(* IEC 61131-3 sources: STAR-PLC-Agent/results/raw/four_group_20261114/star_deepseek_v4/PUB019/generation/sim_00, 1 file *)

(* ---- test_program.st ---- *)
PROGRAM PLC_PRG
VAR
 BenchStep : UDINT := 0;
 BenchCalls : UDINT := 0;
 BenchDone : BOOL := FALSE;
 BenchUut0 : FB_Task;
 BenchUut1 : FB_Task;
 TraceIn_ManualMode : ARRAY[0..12] OF BOOL;
 TraceIn_SingleStepMode : ARRAY[0..12] OF BOOL;
 TraceIn_SingleCycleMode : ARRAY[0..12] OF BOOL;
 TraceIn_ContinuousMode : ARRAY[0..12] OF BOOL;
 TraceIn_EmergencyStop : ARRAY[0..12] OF BOOL;
 TraceIn_Start : ARRAY[0..12] OF BOOL;
 TraceIn_DownButton : ARRAY[0..12] OF BOOL;
 TraceIn_UpButton : ARRAY[0..12] OF BOOL;
 TraceIn_LeftButton : ARRAY[0..12] OF BOOL;
 TraceIn_RightButton : ARRAY[0..12] OF BOOL;
 TraceIn_GripButton : ARRAY[0..12] OF BOOL;
 TraceIn_ReleaseButton : ARRAY[0..12] OF BOOL;
 TraceIn_DownLimitSwitch : ARRAY[0..12] OF BOOL;
 TraceIn_UpLimitSwitch : ARRAY[0..12] OF BOOL;
 TraceIn_LeftLimitSwitch : ARRAY[0..12] OF BOOL;
 TraceIn_RightLimitSwitch : ARRAY[0..12] OF BOOL;
 TraceIn_GripLimitSwitch : ARRAY[0..12] OF BOOL;
 TraceIn_ReleaseLimitSwitch : ARRAY[0..12] OF BOOL;
 TraceOut_MoveDown : ARRAY[0..12] OF BOOL;
 TraceOut_MoveUp : ARRAY[0..12] OF BOOL;
 TraceOut_MoveLeft : ARRAY[0..12] OF BOOL;
 TraceOut_MoveRight : ARRAY[0..12] OF BOOL;
 TraceOut_ActivateGrip : ARRAY[0..12] OF BOOL;
 TraceOut_ActivateRelease : ARRAY[0..12] OF BOOL;
END_VAR

IF NOT BenchDone THEN
 CASE BenchStep OF
 0:
   BenchUut0.ManualMode := TRUE;
   BenchUut0.SingleStepMode := FALSE;
   BenchUut0.SingleCycleMode := FALSE;
   BenchUut0.ContinuousMode := FALSE;
   BenchUut0.EmergencyStop := TRUE;
   BenchUut0.Start := FALSE;
   BenchUut0.DownButton := TRUE;
   BenchUut0.UpButton := FALSE;
   BenchUut0.LeftButton := FALSE;
   BenchUut0.RightButton := FALSE;
   BenchUut0.GripButton := FALSE;
   BenchUut0.ReleaseButton := FALSE;
   BenchUut0.DownLimitSwitch := FALSE;
   BenchUut0.UpLimitSwitch := TRUE;
   BenchUut0.LeftLimitSwitch := TRUE;
   BenchUut0.RightLimitSwitch := FALSE;
   BenchUut0.GripLimitSwitch := FALSE;
   BenchUut0.ReleaseLimitSwitch := FALSE;
   TraceIn_ManualMode[0] := BenchUut0.ManualMode;
   TraceIn_SingleStepMode[0] := BenchUut0.SingleStepMode;
   TraceIn_SingleCycleMode[0] := BenchUut0.SingleCycleMode;
   TraceIn_ContinuousMode[0] := BenchUut0.ContinuousMode;
   TraceIn_EmergencyStop[0] := BenchUut0.EmergencyStop;
   TraceIn_Start[0] := BenchUut0.Start;
   TraceIn_DownButton[0] := BenchUut0.DownButton;
   TraceIn_UpButton[0] := BenchUut0.UpButton;
   TraceIn_LeftButton[0] := BenchUut0.LeftButton;
   TraceIn_RightButton[0] := BenchUut0.RightButton;
   TraceIn_GripButton[0] := BenchUut0.GripButton;
   TraceIn_ReleaseButton[0] := BenchUut0.ReleaseButton;
   TraceIn_DownLimitSwitch[0] := BenchUut0.DownLimitSwitch;
   TraceIn_UpLimitSwitch[0] := BenchUut0.UpLimitSwitch;
   TraceIn_LeftLimitSwitch[0] := BenchUut0.LeftLimitSwitch;
   TraceIn_RightLimitSwitch[0] := BenchUut0.RightLimitSwitch;
   TraceIn_GripLimitSwitch[0] := BenchUut0.GripLimitSwitch;
   TraceIn_ReleaseLimitSwitch[0] := BenchUut0.ReleaseLimitSwitch;
   BenchUut0();
   TraceOut_MoveDown[0] := BenchUut0.MoveDown;
   TraceOut_MoveUp[0] := BenchUut0.MoveUp;
   TraceOut_MoveLeft[0] := BenchUut0.MoveLeft;
   TraceOut_MoveRight[0] := BenchUut0.MoveRight;
   TraceOut_ActivateGrip[0] := BenchUut0.ActivateGrip;
   TraceOut_ActivateRelease[0] := BenchUut0.ActivateRelease;
   BenchCalls := BenchCalls + 1;
 1:
   BenchUut0.ManualMode := TRUE;
   BenchUut0.SingleStepMode := FALSE;
   BenchUut0.SingleCycleMode := FALSE;
   BenchUut0.ContinuousMode := FALSE;
   BenchUut0.EmergencyStop := TRUE;
   BenchUut0.Start := FALSE;
   BenchUut0.DownButton := TRUE;
   BenchUut0.UpButton := FALSE;
   BenchUut0.LeftButton := FALSE;
   BenchUut0.RightButton := FALSE;
   BenchUut0.GripButton := FALSE;
   BenchUut0.ReleaseButton := FALSE;
   BenchUut0.DownLimitSwitch := TRUE;
   BenchUut0.UpLimitSwitch := FALSE;
   BenchUut0.LeftLimitSwitch := TRUE;
   BenchUut0.RightLimitSwitch := FALSE;
   BenchUut0.GripLimitSwitch := FALSE;
   BenchUut0.ReleaseLimitSwitch := FALSE;
   TraceIn_ManualMode[1] := BenchUut0.ManualMode;
   TraceIn_SingleStepMode[1] := BenchUut0.SingleStepMode;
   TraceIn_SingleCycleMode[1] := BenchUut0.SingleCycleMode;
   TraceIn_ContinuousMode[1] := BenchUut0.ContinuousMode;
   TraceIn_EmergencyStop[1] := BenchUut0.EmergencyStop;
   TraceIn_Start[1] := BenchUut0.Start;
   TraceIn_DownButton[1] := BenchUut0.DownButton;
   TraceIn_UpButton[1] := BenchUut0.UpButton;
   TraceIn_LeftButton[1] := BenchUut0.LeftButton;
   TraceIn_RightButton[1] := BenchUut0.RightButton;
   TraceIn_GripButton[1] := BenchUut0.GripButton;
   TraceIn_ReleaseButton[1] := BenchUut0.ReleaseButton;
   TraceIn_DownLimitSwitch[1] := BenchUut0.DownLimitSwitch;
   TraceIn_UpLimitSwitch[1] := BenchUut0.UpLimitSwitch;
   TraceIn_LeftLimitSwitch[1] := BenchUut0.LeftLimitSwitch;
   TraceIn_RightLimitSwitch[1] := BenchUut0.RightLimitSwitch;
   TraceIn_GripLimitSwitch[1] := BenchUut0.GripLimitSwitch;
   TraceIn_ReleaseLimitSwitch[1] := BenchUut0.ReleaseLimitSwitch;
   BenchUut0();
   TraceOut_MoveDown[1] := BenchUut0.MoveDown;
   TraceOut_MoveUp[1] := BenchUut0.MoveUp;
   TraceOut_MoveLeft[1] := BenchUut0.MoveLeft;
   TraceOut_MoveRight[1] := BenchUut0.MoveRight;
   TraceOut_ActivateGrip[1] := BenchUut0.ActivateGrip;
   TraceOut_ActivateRelease[1] := BenchUut0.ActivateRelease;
   BenchCalls := BenchCalls + 1;
 2:
   BenchUut0.ManualMode := TRUE;
   BenchUut0.SingleStepMode := FALSE;
   BenchUut0.SingleCycleMode := FALSE;
   BenchUut0.ContinuousMode := FALSE;
   BenchUut0.EmergencyStop := FALSE;
   BenchUut0.Start := FALSE;
   BenchUut0.DownButton := TRUE;
   BenchUut0.UpButton := FALSE;
   BenchUut0.LeftButton := FALSE;
   BenchUut0.RightButton := FALSE;
   BenchUut0.GripButton := FALSE;
   BenchUut0.ReleaseButton := FALSE;
   BenchUut0.DownLimitSwitch := FALSE;
   BenchUut0.UpLimitSwitch := TRUE;
   BenchUut0.LeftLimitSwitch := TRUE;
   BenchUut0.RightLimitSwitch := FALSE;
   BenchUut0.GripLimitSwitch := FALSE;
   BenchUut0.ReleaseLimitSwitch := FALSE;
   TraceIn_ManualMode[2] := BenchUut0.ManualMode;
   TraceIn_SingleStepMode[2] := BenchUut0.SingleStepMode;
   TraceIn_SingleCycleMode[2] := BenchUut0.SingleCycleMode;
   TraceIn_ContinuousMode[2] := BenchUut0.ContinuousMode;
   TraceIn_EmergencyStop[2] := BenchUut0.EmergencyStop;
   TraceIn_Start[2] := BenchUut0.Start;
   TraceIn_DownButton[2] := BenchUut0.DownButton;
   TraceIn_UpButton[2] := BenchUut0.UpButton;
   TraceIn_LeftButton[2] := BenchUut0.LeftButton;
   TraceIn_RightButton[2] := BenchUut0.RightButton;
   TraceIn_GripButton[2] := BenchUut0.GripButton;
   TraceIn_ReleaseButton[2] := BenchUut0.ReleaseButton;
   TraceIn_DownLimitSwitch[2] := BenchUut0.DownLimitSwitch;
   TraceIn_UpLimitSwitch[2] := BenchUut0.UpLimitSwitch;
   TraceIn_LeftLimitSwitch[2] := BenchUut0.LeftLimitSwitch;
   TraceIn_RightLimitSwitch[2] := BenchUut0.RightLimitSwitch;
   TraceIn_GripLimitSwitch[2] := BenchUut0.GripLimitSwitch;
   TraceIn_ReleaseLimitSwitch[2] := BenchUut0.ReleaseLimitSwitch;
   BenchUut0();
   TraceOut_MoveDown[2] := BenchUut0.MoveDown;
   TraceOut_MoveUp[2] := BenchUut0.MoveUp;
   TraceOut_MoveLeft[2] := BenchUut0.MoveLeft;
   TraceOut_MoveRight[2] := BenchUut0.MoveRight;
   TraceOut_ActivateGrip[2] := BenchUut0.ActivateGrip;
   TraceOut_ActivateRelease[2] := BenchUut0.ActivateRelease;
   BenchCalls := BenchCalls + 1;
 3:
   BenchUut0.ManualMode := TRUE;
   BenchUut0.SingleStepMode := FALSE;
   BenchUut0.SingleCycleMode := FALSE;
   BenchUut0.ContinuousMode := FALSE;
   BenchUut0.EmergencyStop := TRUE;
   BenchUut0.Start := FALSE;
   BenchUut0.DownButton := TRUE;
   BenchUut0.UpButton := FALSE;
   BenchUut0.LeftButton := FALSE;
   BenchUut0.RightButton := FALSE;
   BenchUut0.GripButton := FALSE;
   BenchUut0.ReleaseButton := FALSE;
   BenchUut0.DownLimitSwitch := FALSE;
   BenchUut0.UpLimitSwitch := TRUE;
   BenchUut0.LeftLimitSwitch := TRUE;
   BenchUut0.RightLimitSwitch := FALSE;
   BenchUut0.GripLimitSwitch := FALSE;
   BenchUut0.ReleaseLimitSwitch := FALSE;
   TraceIn_ManualMode[3] := BenchUut0.ManualMode;
   TraceIn_SingleStepMode[3] := BenchUut0.SingleStepMode;
   TraceIn_SingleCycleMode[3] := BenchUut0.SingleCycleMode;
   TraceIn_ContinuousMode[3] := BenchUut0.ContinuousMode;
   TraceIn_EmergencyStop[3] := BenchUut0.EmergencyStop;
   TraceIn_Start[3] := BenchUut0.Start;
   TraceIn_DownButton[3] := BenchUut0.DownButton;
   TraceIn_UpButton[3] := BenchUut0.UpButton;
   TraceIn_LeftButton[3] := BenchUut0.LeftButton;
   TraceIn_RightButton[3] := BenchUut0.RightButton;
   TraceIn_GripButton[3] := BenchUut0.GripButton;
   TraceIn_ReleaseButton[3] := BenchUut0.ReleaseButton;
   TraceIn_DownLimitSwitch[3] := BenchUut0.DownLimitSwitch;
   TraceIn_UpLimitSwitch[3] := BenchUut0.UpLimitSwitch;
   TraceIn_LeftLimitSwitch[3] := BenchUut0.LeftLimitSwitch;
   TraceIn_RightLimitSwitch[3] := BenchUut0.RightLimitSwitch;
   TraceIn_GripLimitSwitch[3] := BenchUut0.GripLimitSwitch;
   TraceIn_ReleaseLimitSwitch[3] := BenchUut0.ReleaseLimitSwitch;
   BenchUut0();
   TraceOut_MoveDown[3] := BenchUut0.MoveDown;
   TraceOut_MoveUp[3] := BenchUut0.MoveUp;
   TraceOut_MoveLeft[3] := BenchUut0.MoveLeft;
   TraceOut_MoveRight[3] := BenchUut0.MoveRight;
   TraceOut_ActivateGrip[3] := BenchUut0.ActivateGrip;
   TraceOut_ActivateRelease[3] := BenchUut0.ActivateRelease;
   BenchCalls := BenchCalls + 1;
 4:
   BenchUut0.ManualMode := TRUE;
   BenchUut0.SingleStepMode := FALSE;
   BenchUut0.SingleCycleMode := FALSE;
   BenchUut0.ContinuousMode := FALSE;
   BenchUut0.EmergencyStop := TRUE;
   BenchUut0.Start := FALSE;
   BenchUut0.DownButton := TRUE;
   BenchUut0.UpButton := TRUE;
   BenchUut0.LeftButton := FALSE;
   BenchUut0.RightButton := FALSE;
   BenchUut0.GripButton := FALSE;
   BenchUut0.ReleaseButton := FALSE;
   BenchUut0.DownLimitSwitch := FALSE;
   BenchUut0.UpLimitSwitch := FALSE;
   BenchUut0.LeftLimitSwitch := TRUE;
   BenchUut0.RightLimitSwitch := FALSE;
   BenchUut0.GripLimitSwitch := FALSE;
   BenchUut0.ReleaseLimitSwitch := FALSE;
   TraceIn_ManualMode[4] := BenchUut0.ManualMode;
   TraceIn_SingleStepMode[4] := BenchUut0.SingleStepMode;
   TraceIn_SingleCycleMode[4] := BenchUut0.SingleCycleMode;
   TraceIn_ContinuousMode[4] := BenchUut0.ContinuousMode;
   TraceIn_EmergencyStop[4] := BenchUut0.EmergencyStop;
   TraceIn_Start[4] := BenchUut0.Start;
   TraceIn_DownButton[4] := BenchUut0.DownButton;
   TraceIn_UpButton[4] := BenchUut0.UpButton;
   TraceIn_LeftButton[4] := BenchUut0.LeftButton;
   TraceIn_RightButton[4] := BenchUut0.RightButton;
   TraceIn_GripButton[4] := BenchUut0.GripButton;
   TraceIn_ReleaseButton[4] := BenchUut0.ReleaseButton;
   TraceIn_DownLimitSwitch[4] := BenchUut0.DownLimitSwitch;
   TraceIn_UpLimitSwitch[4] := BenchUut0.UpLimitSwitch;
   TraceIn_LeftLimitSwitch[4] := BenchUut0.LeftLimitSwitch;
   TraceIn_RightLimitSwitch[4] := BenchUut0.RightLimitSwitch;
   TraceIn_GripLimitSwitch[4] := BenchUut0.GripLimitSwitch;
   TraceIn_ReleaseLimitSwitch[4] := BenchUut0.ReleaseLimitSwitch;
   BenchUut0();
   TraceOut_MoveDown[4] := BenchUut0.MoveDown;
   TraceOut_MoveUp[4] := BenchUut0.MoveUp;
   TraceOut_MoveLeft[4] := BenchUut0.MoveLeft;
   TraceOut_MoveRight[4] := BenchUut0.MoveRight;
   TraceOut_ActivateGrip[4] := BenchUut0.ActivateGrip;
   TraceOut_ActivateRelease[4] := BenchUut0.ActivateRelease;
   BenchCalls := BenchCalls + 1;
 5:
   BenchUut1.ManualMode := FALSE;
   BenchUut1.SingleStepMode := FALSE;
   BenchUut1.SingleCycleMode := TRUE;
   BenchUut1.ContinuousMode := FALSE;
   BenchUut1.EmergencyStop := TRUE;
   BenchUut1.Start := TRUE;
   BenchUut1.DownButton := FALSE;
   BenchUut1.UpButton := FALSE;
   BenchUut1.LeftButton := FALSE;
   BenchUut1.RightButton := FALSE;
   BenchUut1.GripButton := FALSE;
   BenchUut1.ReleaseButton := FALSE;
   BenchUut1.DownLimitSwitch := FALSE;
   BenchUut1.UpLimitSwitch := TRUE;
   BenchUut1.LeftLimitSwitch := TRUE;
   BenchUut1.RightLimitSwitch := FALSE;
   BenchUut1.GripLimitSwitch := FALSE;
   BenchUut1.ReleaseLimitSwitch := FALSE;
   TraceIn_ManualMode[5] := BenchUut1.ManualMode;
   TraceIn_SingleStepMode[5] := BenchUut1.SingleStepMode;
   TraceIn_SingleCycleMode[5] := BenchUut1.SingleCycleMode;
   TraceIn_ContinuousMode[5] := BenchUut1.ContinuousMode;
   TraceIn_EmergencyStop[5] := BenchUut1.EmergencyStop;
   TraceIn_Start[5] := BenchUut1.Start;
   TraceIn_DownButton[5] := BenchUut1.DownButton;
   TraceIn_UpButton[5] := BenchUut1.UpButton;
   TraceIn_LeftButton[5] := BenchUut1.LeftButton;
   TraceIn_RightButton[5] := BenchUut1.RightButton;
   TraceIn_GripButton[5] := BenchUut1.GripButton;
   TraceIn_ReleaseButton[5] := BenchUut1.ReleaseButton;
   TraceIn_DownLimitSwitch[5] := BenchUut1.DownLimitSwitch;
   TraceIn_UpLimitSwitch[5] := BenchUut1.UpLimitSwitch;
   TraceIn_LeftLimitSwitch[5] := BenchUut1.LeftLimitSwitch;
   TraceIn_RightLimitSwitch[5] := BenchUut1.RightLimitSwitch;
   TraceIn_GripLimitSwitch[5] := BenchUut1.GripLimitSwitch;
   TraceIn_ReleaseLimitSwitch[5] := BenchUut1.ReleaseLimitSwitch;
   BenchUut1();
   TraceOut_MoveDown[5] := BenchUut1.MoveDown;
   TraceOut_MoveUp[5] := BenchUut1.MoveUp;
   TraceOut_MoveLeft[5] := BenchUut1.MoveLeft;
   TraceOut_MoveRight[5] := BenchUut1.MoveRight;
   TraceOut_ActivateGrip[5] := BenchUut1.ActivateGrip;
   TraceOut_ActivateRelease[5] := BenchUut1.ActivateRelease;
   BenchCalls := BenchCalls + 1;
 6:
   BenchUut1.ManualMode := FALSE;
   BenchUut1.SingleStepMode := FALSE;
   BenchUut1.SingleCycleMode := TRUE;
   BenchUut1.ContinuousMode := FALSE;
   BenchUut1.EmergencyStop := TRUE;
   BenchUut1.Start := FALSE;
   BenchUut1.DownButton := FALSE;
   BenchUut1.UpButton := FALSE;
   BenchUut1.LeftButton := FALSE;
   BenchUut1.RightButton := FALSE;
   BenchUut1.GripButton := FALSE;
   BenchUut1.ReleaseButton := FALSE;
   BenchUut1.DownLimitSwitch := TRUE;
   BenchUut1.UpLimitSwitch := FALSE;
   BenchUut1.LeftLimitSwitch := TRUE;
   BenchUut1.RightLimitSwitch := FALSE;
   BenchUut1.GripLimitSwitch := FALSE;
   BenchUut1.ReleaseLimitSwitch := FALSE;
   TraceIn_ManualMode[6] := BenchUut1.ManualMode;
   TraceIn_SingleStepMode[6] := BenchUut1.SingleStepMode;
   TraceIn_SingleCycleMode[6] := BenchUut1.SingleCycleMode;
   TraceIn_ContinuousMode[6] := BenchUut1.ContinuousMode;
   TraceIn_EmergencyStop[6] := BenchUut1.EmergencyStop;
   TraceIn_Start[6] := BenchUut1.Start;
   TraceIn_DownButton[6] := BenchUut1.DownButton;
   TraceIn_UpButton[6] := BenchUut1.UpButton;
   TraceIn_LeftButton[6] := BenchUut1.LeftButton;
   TraceIn_RightButton[6] := BenchUut1.RightButton;
   TraceIn_GripButton[6] := BenchUut1.GripButton;
   TraceIn_ReleaseButton[6] := BenchUut1.ReleaseButton;
   TraceIn_DownLimitSwitch[6] := BenchUut1.DownLimitSwitch;
   TraceIn_UpLimitSwitch[6] := BenchUut1.UpLimitSwitch;
   TraceIn_LeftLimitSwitch[6] := BenchUut1.LeftLimitSwitch;
   TraceIn_RightLimitSwitch[6] := BenchUut1.RightLimitSwitch;
   TraceIn_GripLimitSwitch[6] := BenchUut1.GripLimitSwitch;
   TraceIn_ReleaseLimitSwitch[6] := BenchUut1.ReleaseLimitSwitch;
   BenchUut1();
   TraceOut_MoveDown[6] := BenchUut1.MoveDown;
   TraceOut_MoveUp[6] := BenchUut1.MoveUp;
   TraceOut_MoveLeft[6] := BenchUut1.MoveLeft;
   TraceOut_MoveRight[6] := BenchUut1.MoveRight;
   TraceOut_ActivateGrip[6] := BenchUut1.ActivateGrip;
   TraceOut_ActivateRelease[6] := BenchUut1.ActivateRelease;
   BenchCalls := BenchCalls + 1;
 7:
   BenchUut1.ManualMode := FALSE;
   BenchUut1.SingleStepMode := FALSE;
   BenchUut1.SingleCycleMode := TRUE;
   BenchUut1.ContinuousMode := FALSE;
   BenchUut1.EmergencyStop := TRUE;
   BenchUut1.Start := FALSE;
   BenchUut1.DownButton := FALSE;
   BenchUut1.UpButton := FALSE;
   BenchUut1.LeftButton := FALSE;
   BenchUut1.RightButton := FALSE;
   BenchUut1.GripButton := FALSE;
   BenchUut1.ReleaseButton := FALSE;
   BenchUut1.DownLimitSwitch := TRUE;
   BenchUut1.UpLimitSwitch := FALSE;
   BenchUut1.LeftLimitSwitch := TRUE;
   BenchUut1.RightLimitSwitch := FALSE;
   BenchUut1.GripLimitSwitch := TRUE;
   BenchUut1.ReleaseLimitSwitch := FALSE;
   TraceIn_ManualMode[7] := BenchUut1.ManualMode;
   TraceIn_SingleStepMode[7] := BenchUut1.SingleStepMode;
   TraceIn_SingleCycleMode[7] := BenchUut1.SingleCycleMode;
   TraceIn_ContinuousMode[7] := BenchUut1.ContinuousMode;
   TraceIn_EmergencyStop[7] := BenchUut1.EmergencyStop;
   TraceIn_Start[7] := BenchUut1.Start;
   TraceIn_DownButton[7] := BenchUut1.DownButton;
   TraceIn_UpButton[7] := BenchUut1.UpButton;
   TraceIn_LeftButton[7] := BenchUut1.LeftButton;
   TraceIn_RightButton[7] := BenchUut1.RightButton;
   TraceIn_GripButton[7] := BenchUut1.GripButton;
   TraceIn_ReleaseButton[7] := BenchUut1.ReleaseButton;
   TraceIn_DownLimitSwitch[7] := BenchUut1.DownLimitSwitch;
   TraceIn_UpLimitSwitch[7] := BenchUut1.UpLimitSwitch;
   TraceIn_LeftLimitSwitch[7] := BenchUut1.LeftLimitSwitch;
   TraceIn_RightLimitSwitch[7] := BenchUut1.RightLimitSwitch;
   TraceIn_GripLimitSwitch[7] := BenchUut1.GripLimitSwitch;
   TraceIn_ReleaseLimitSwitch[7] := BenchUut1.ReleaseLimitSwitch;
   BenchUut1();
   TraceOut_MoveDown[7] := BenchUut1.MoveDown;
   TraceOut_MoveUp[7] := BenchUut1.MoveUp;
   TraceOut_MoveLeft[7] := BenchUut1.MoveLeft;
   TraceOut_MoveRight[7] := BenchUut1.MoveRight;
   TraceOut_ActivateGrip[7] := BenchUut1.ActivateGrip;
   TraceOut_ActivateRelease[7] := BenchUut1.ActivateRelease;
   BenchCalls := BenchCalls + 1;
 8:
   BenchUut1.ManualMode := FALSE;
   BenchUut1.SingleStepMode := FALSE;
   BenchUut1.SingleCycleMode := TRUE;
   BenchUut1.ContinuousMode := FALSE;
   BenchUut1.EmergencyStop := TRUE;
   BenchUut1.Start := FALSE;
   BenchUut1.DownButton := FALSE;
   BenchUut1.UpButton := FALSE;
   BenchUut1.LeftButton := FALSE;
   BenchUut1.RightButton := FALSE;
   BenchUut1.GripButton := FALSE;
   BenchUut1.ReleaseButton := FALSE;
   BenchUut1.DownLimitSwitch := FALSE;
   BenchUut1.UpLimitSwitch := TRUE;
   BenchUut1.LeftLimitSwitch := TRUE;
   BenchUut1.RightLimitSwitch := FALSE;
   BenchUut1.GripLimitSwitch := TRUE;
   BenchUut1.ReleaseLimitSwitch := FALSE;
   TraceIn_ManualMode[8] := BenchUut1.ManualMode;
   TraceIn_SingleStepMode[8] := BenchUut1.SingleStepMode;
   TraceIn_SingleCycleMode[8] := BenchUut1.SingleCycleMode;
   TraceIn_ContinuousMode[8] := BenchUut1.ContinuousMode;
   TraceIn_EmergencyStop[8] := BenchUut1.EmergencyStop;
   TraceIn_Start[8] := BenchUut1.Start;
   TraceIn_DownButton[8] := BenchUut1.DownButton;
   TraceIn_UpButton[8] := BenchUut1.UpButton;
   TraceIn_LeftButton[8] := BenchUut1.LeftButton;
   TraceIn_RightButton[8] := BenchUut1.RightButton;
   TraceIn_GripButton[8] := BenchUut1.GripButton;
   TraceIn_ReleaseButton[8] := BenchUut1.ReleaseButton;
   TraceIn_DownLimitSwitch[8] := BenchUut1.DownLimitSwitch;
   TraceIn_UpLimitSwitch[8] := BenchUut1.UpLimitSwitch;
   TraceIn_LeftLimitSwitch[8] := BenchUut1.LeftLimitSwitch;
   TraceIn_RightLimitSwitch[8] := BenchUut1.RightLimitSwitch;
   TraceIn_GripLimitSwitch[8] := BenchUut1.GripLimitSwitch;
   TraceIn_ReleaseLimitSwitch[8] := BenchUut1.ReleaseLimitSwitch;
   BenchUut1();
   TraceOut_MoveDown[8] := BenchUut1.MoveDown;
   TraceOut_MoveUp[8] := BenchUut1.MoveUp;
   TraceOut_MoveLeft[8] := BenchUut1.MoveLeft;
   TraceOut_MoveRight[8] := BenchUut1.MoveRight;
   TraceOut_ActivateGrip[8] := BenchUut1.ActivateGrip;
   TraceOut_ActivateRelease[8] := BenchUut1.ActivateRelease;
   BenchCalls := BenchCalls + 1;
 9:
   BenchUut1.ManualMode := FALSE;
   BenchUut1.SingleStepMode := FALSE;
   BenchUut1.SingleCycleMode := TRUE;
   BenchUut1.ContinuousMode := FALSE;
   BenchUut1.EmergencyStop := TRUE;
   BenchUut1.Start := FALSE;
   BenchUut1.DownButton := FALSE;
   BenchUut1.UpButton := FALSE;
   BenchUut1.LeftButton := FALSE;
   BenchUut1.RightButton := FALSE;
   BenchUut1.GripButton := FALSE;
   BenchUut1.ReleaseButton := FALSE;
   BenchUut1.DownLimitSwitch := FALSE;
   BenchUut1.UpLimitSwitch := TRUE;
   BenchUut1.LeftLimitSwitch := FALSE;
   BenchUut1.RightLimitSwitch := TRUE;
   BenchUut1.GripLimitSwitch := TRUE;
   BenchUut1.ReleaseLimitSwitch := FALSE;
   TraceIn_ManualMode[9] := BenchUut1.ManualMode;
   TraceIn_SingleStepMode[9] := BenchUut1.SingleStepMode;
   TraceIn_SingleCycleMode[9] := BenchUut1.SingleCycleMode;
   TraceIn_ContinuousMode[9] := BenchUut1.ContinuousMode;
   TraceIn_EmergencyStop[9] := BenchUut1.EmergencyStop;
   TraceIn_Start[9] := BenchUut1.Start;
   TraceIn_DownButton[9] := BenchUut1.DownButton;
   TraceIn_UpButton[9] := BenchUut1.UpButton;
   TraceIn_LeftButton[9] := BenchUut1.LeftButton;
   TraceIn_RightButton[9] := BenchUut1.RightButton;
   TraceIn_GripButton[9] := BenchUut1.GripButton;
   TraceIn_ReleaseButton[9] := BenchUut1.ReleaseButton;
   TraceIn_DownLimitSwitch[9] := BenchUut1.DownLimitSwitch;
   TraceIn_UpLimitSwitch[9] := BenchUut1.UpLimitSwitch;
   TraceIn_LeftLimitSwitch[9] := BenchUut1.LeftLimitSwitch;
   TraceIn_RightLimitSwitch[9] := BenchUut1.RightLimitSwitch;
   TraceIn_GripLimitSwitch[9] := BenchUut1.GripLimitSwitch;
   TraceIn_ReleaseLimitSwitch[9] := BenchUut1.ReleaseLimitSwitch;
   BenchUut1();
   TraceOut_MoveDown[9] := BenchUut1.MoveDown;
   TraceOut_MoveUp[9] := BenchUut1.MoveUp;
   TraceOut_MoveLeft[9] := BenchUut1.MoveLeft;
   TraceOut_MoveRight[9] := BenchUut1.MoveRight;
   TraceOut_ActivateGrip[9] := BenchUut1.ActivateGrip;
   TraceOut_ActivateRelease[9] := BenchUut1.ActivateRelease;
   BenchCalls := BenchCalls + 1;
 10:
   BenchUut1.ManualMode := FALSE;
   BenchUut1.SingleStepMode := FALSE;
   BenchUut1.SingleCycleMode := TRUE;
   BenchUut1.ContinuousMode := FALSE;
   BenchUut1.EmergencyStop := TRUE;
   BenchUut1.Start := FALSE;
   BenchUut1.DownButton := FALSE;
   BenchUut1.UpButton := FALSE;
   BenchUut1.LeftButton := FALSE;
   BenchUut1.RightButton := FALSE;
   BenchUut1.GripButton := FALSE;
   BenchUut1.ReleaseButton := FALSE;
   BenchUut1.DownLimitSwitch := TRUE;
   BenchUut1.UpLimitSwitch := FALSE;
   BenchUut1.LeftLimitSwitch := FALSE;
   BenchUut1.RightLimitSwitch := TRUE;
   BenchUut1.GripLimitSwitch := TRUE;
   BenchUut1.ReleaseLimitSwitch := FALSE;
   TraceIn_ManualMode[10] := BenchUut1.ManualMode;
   TraceIn_SingleStepMode[10] := BenchUut1.SingleStepMode;
   TraceIn_SingleCycleMode[10] := BenchUut1.SingleCycleMode;
   TraceIn_ContinuousMode[10] := BenchUut1.ContinuousMode;
   TraceIn_EmergencyStop[10] := BenchUut1.EmergencyStop;
   TraceIn_Start[10] := BenchUut1.Start;
   TraceIn_DownButton[10] := BenchUut1.DownButton;
   TraceIn_UpButton[10] := BenchUut1.UpButton;
   TraceIn_LeftButton[10] := BenchUut1.LeftButton;
   TraceIn_RightButton[10] := BenchUut1.RightButton;
   TraceIn_GripButton[10] := BenchUut1.GripButton;
   TraceIn_ReleaseButton[10] := BenchUut1.ReleaseButton;
   TraceIn_DownLimitSwitch[10] := BenchUut1.DownLimitSwitch;
   TraceIn_UpLimitSwitch[10] := BenchUut1.UpLimitSwitch;
   TraceIn_LeftLimitSwitch[10] := BenchUut1.LeftLimitSwitch;
   TraceIn_RightLimitSwitch[10] := BenchUut1.RightLimitSwitch;
   TraceIn_GripLimitSwitch[10] := BenchUut1.GripLimitSwitch;
   TraceIn_ReleaseLimitSwitch[10] := BenchUut1.ReleaseLimitSwitch;
   BenchUut1();
   TraceOut_MoveDown[10] := BenchUut1.MoveDown;
   TraceOut_MoveUp[10] := BenchUut1.MoveUp;
   TraceOut_MoveLeft[10] := BenchUut1.MoveLeft;
   TraceOut_MoveRight[10] := BenchUut1.MoveRight;
   TraceOut_ActivateGrip[10] := BenchUut1.ActivateGrip;
   TraceOut_ActivateRelease[10] := BenchUut1.ActivateRelease;
   BenchCalls := BenchCalls + 1;
 11:
   BenchUut1.ManualMode := FALSE;
   BenchUut1.SingleStepMode := FALSE;
   BenchUut1.SingleCycleMode := TRUE;
   BenchUut1.ContinuousMode := FALSE;
   BenchUut1.EmergencyStop := TRUE;
   BenchUut1.Start := FALSE;
   BenchUut1.DownButton := FALSE;
   BenchUut1.UpButton := FALSE;
   BenchUut1.LeftButton := FALSE;
   BenchUut1.RightButton := FALSE;
   BenchUut1.GripButton := FALSE;
   BenchUut1.ReleaseButton := FALSE;
   BenchUut1.DownLimitSwitch := TRUE;
   BenchUut1.UpLimitSwitch := FALSE;
   BenchUut1.LeftLimitSwitch := FALSE;
   BenchUut1.RightLimitSwitch := TRUE;
   BenchUut1.GripLimitSwitch := FALSE;
   BenchUut1.ReleaseLimitSwitch := TRUE;
   TraceIn_ManualMode[11] := BenchUut1.ManualMode;
   TraceIn_SingleStepMode[11] := BenchUut1.SingleStepMode;
   TraceIn_SingleCycleMode[11] := BenchUut1.SingleCycleMode;
   TraceIn_ContinuousMode[11] := BenchUut1.ContinuousMode;
   TraceIn_EmergencyStop[11] := BenchUut1.EmergencyStop;
   TraceIn_Start[11] := BenchUut1.Start;
   TraceIn_DownButton[11] := BenchUut1.DownButton;
   TraceIn_UpButton[11] := BenchUut1.UpButton;
   TraceIn_LeftButton[11] := BenchUut1.LeftButton;
   TraceIn_RightButton[11] := BenchUut1.RightButton;
   TraceIn_GripButton[11] := BenchUut1.GripButton;
   TraceIn_ReleaseButton[11] := BenchUut1.ReleaseButton;
   TraceIn_DownLimitSwitch[11] := BenchUut1.DownLimitSwitch;
   TraceIn_UpLimitSwitch[11] := BenchUut1.UpLimitSwitch;
   TraceIn_LeftLimitSwitch[11] := BenchUut1.LeftLimitSwitch;
   TraceIn_RightLimitSwitch[11] := BenchUut1.RightLimitSwitch;
   TraceIn_GripLimitSwitch[11] := BenchUut1.GripLimitSwitch;
   TraceIn_ReleaseLimitSwitch[11] := BenchUut1.ReleaseLimitSwitch;
   BenchUut1();
   TraceOut_MoveDown[11] := BenchUut1.MoveDown;
   TraceOut_MoveUp[11] := BenchUut1.MoveUp;
   TraceOut_MoveLeft[11] := BenchUut1.MoveLeft;
   TraceOut_MoveRight[11] := BenchUut1.MoveRight;
   TraceOut_ActivateGrip[11] := BenchUut1.ActivateGrip;
   TraceOut_ActivateRelease[11] := BenchUut1.ActivateRelease;
   BenchCalls := BenchCalls + 1;
 12:
   BenchUut1.ManualMode := FALSE;
   BenchUut1.SingleStepMode := FALSE;
   BenchUut1.SingleCycleMode := TRUE;
   BenchUut1.ContinuousMode := FALSE;
   BenchUut1.EmergencyStop := TRUE;
   BenchUut1.Start := FALSE;
   BenchUut1.DownButton := FALSE;
   BenchUut1.UpButton := FALSE;
   BenchUut1.LeftButton := FALSE;
   BenchUut1.RightButton := FALSE;
   BenchUut1.GripButton := FALSE;
   BenchUut1.ReleaseButton := FALSE;
   BenchUut1.DownLimitSwitch := FALSE;
   BenchUut1.UpLimitSwitch := TRUE;
   BenchUut1.LeftLimitSwitch := FALSE;
   BenchUut1.RightLimitSwitch := TRUE;
   BenchUut1.GripLimitSwitch := FALSE;
   BenchUut1.ReleaseLimitSwitch := TRUE;
   TraceIn_ManualMode[12] := BenchUut1.ManualMode;
   TraceIn_SingleStepMode[12] := BenchUut1.SingleStepMode;
   TraceIn_SingleCycleMode[12] := BenchUut1.SingleCycleMode;
   TraceIn_ContinuousMode[12] := BenchUut1.ContinuousMode;
   TraceIn_EmergencyStop[12] := BenchUut1.EmergencyStop;
   TraceIn_Start[12] := BenchUut1.Start;
   TraceIn_DownButton[12] := BenchUut1.DownButton;
   TraceIn_UpButton[12] := BenchUut1.UpButton;
   TraceIn_LeftButton[12] := BenchUut1.LeftButton;
   TraceIn_RightButton[12] := BenchUut1.RightButton;
   TraceIn_GripButton[12] := BenchUut1.GripButton;
   TraceIn_ReleaseButton[12] := BenchUut1.ReleaseButton;
   TraceIn_DownLimitSwitch[12] := BenchUut1.DownLimitSwitch;
   TraceIn_UpLimitSwitch[12] := BenchUut1.UpLimitSwitch;
   TraceIn_LeftLimitSwitch[12] := BenchUut1.LeftLimitSwitch;
   TraceIn_RightLimitSwitch[12] := BenchUut1.RightLimitSwitch;
   TraceIn_GripLimitSwitch[12] := BenchUut1.GripLimitSwitch;
   TraceIn_ReleaseLimitSwitch[12] := BenchUut1.ReleaseLimitSwitch;
   BenchUut1();
   TraceOut_MoveDown[12] := BenchUut1.MoveDown;
   TraceOut_MoveUp[12] := BenchUut1.MoveUp;
   TraceOut_MoveLeft[12] := BenchUut1.MoveLeft;
   TraceOut_MoveRight[12] := BenchUut1.MoveRight;
   TraceOut_ActivateGrip[12] := BenchUut1.ActivateGrip;
   TraceOut_ActivateRelease[12] := BenchUut1.ActivateRelease;
   BenchCalls := BenchCalls + 1;
 END_CASE;
 BenchStep := BenchStep + 1;
 IF BenchStep >= 13 THEN BenchDone := TRUE; END_IF;
END_IF;
END_PROGRAM
